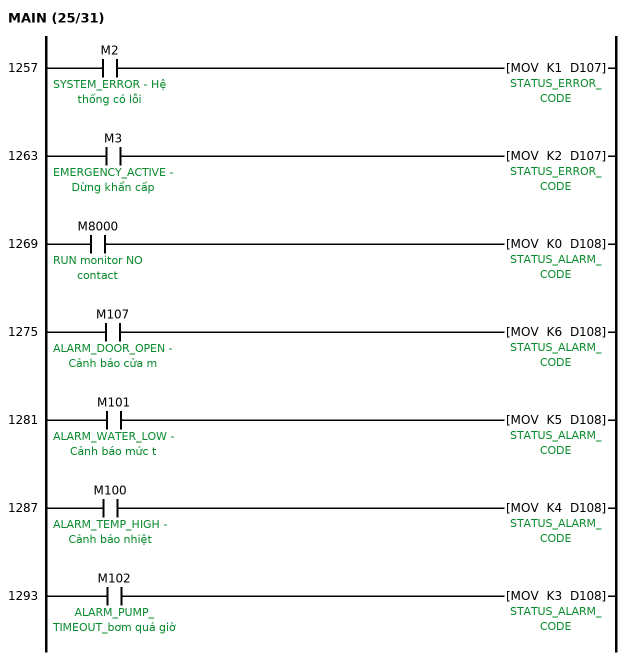
[picture p24: ladder of MAIN, rungs at steps 1257 to 1293]
1257  LD      M2  ; SYSTEM_ERROR - Hệ thống có lỗi
      MOV     K1 D107
1263  LD      M3  ; EMERGENCY_ACTIVE - Dừng khẩn cấp
      MOV     K2 D107
1269  LD      M8000  ; RUN monitor NO contact
      MOV     K0 D108  ; STATUS_ALARM_CODE
1275  LD      M107  ; ALARM_DOOR_OPEN - Cảnh báo cửa m
      MOV     K6 D108
1281  LD      M101  ; ALARM_WATER_LOW - Cảnh báo mức t
      MOV     K5 D108
1287  LD      M100  ; ALARM_TEMP_HIGH - Cảnh báo nhiệt
      MOV     K4 D108
1293  LD      M102  ; ALARM_PUMP_TIMEOUT_bơm quá giờ
      MOV     K3 D108
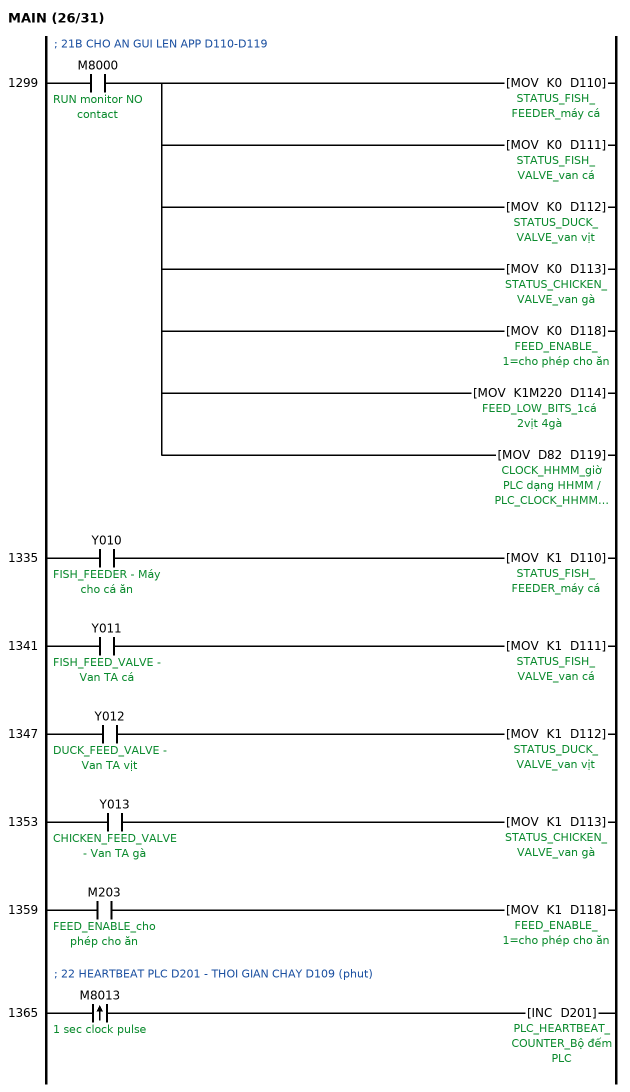
; 21B CHO AN GUI LEN APP D110-D119
1299  LD      M8000  ; RUN monitor NO contact
      MOV     K0 D110  ; STATUS_FISH_FEEDER_máy cá
      MOV     K0 D111  ; STATUS_FISH_VALVE_van cá
      MOV     K0 D112  ; STATUS_DUCK_VALVE_van vịt
      MOV     K0 D113  ; STATUS_CHICKEN_VALVE_van gà
      MOV     K0 D118  ; FEED_ENABLE_1=cho phép cho ăn
      MOV     K1M220 D114  ; FEED_LOW_BITS_1cá 2vịt 4gà
      MOV     D82 D119  ; PLC_CLOCK_HHMM_giờ PLC
1335  LD      Y010  ; FISH_FEEDER - Máy cho cá ăn
      MOV     K1 D110
1341  LD      Y011  ; FISH_FEED_VALVE - Van TA cá
      MOV     K1 D111
1347  LD      Y012  ; DUCK_FEED_VALVE - Van TA vịt
      MOV     K1 D112
1353  LD      Y013  ; CHICKEN_FEED_VALVE - Van TA gà
      MOV     K1 D113
1359  LD      M203  ; FEED_ENABLE_cho phép cho ăn
      MOV     K1 D118
; 22 HEARTBEAT PLC D201 - THOI GIAN CHAY D109 (phut)
1365  LDP     M8013  ; 1 sec clock pulse
      INC     D201  ; PLC_HEARTBEAT_COUNTER_Bộ đếm PLC
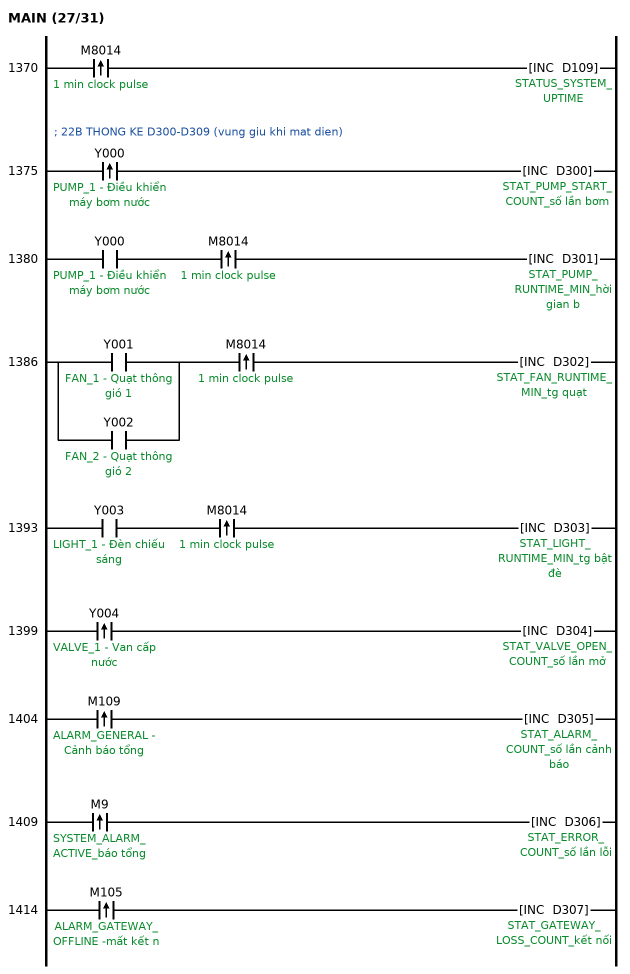
1370  LDP     M8014  ; 1 min clock pulse
      INC     D109  ; STATUS_SYSTEM_UPTIME
; 22B THONG KE D300-D309 (vung giu khi mat dien)
1375  LDP     Y000  ; PUMP_1 - Điều khiển máy bơm nước
      INC     D300  ; STAT_PUMP_START_COUNT_số lần bơm
1380  LD      Y000  ; PUMP_1 - Điều khiển máy bơm nước
      ANDP    M8014  ; 1 min clock pulse
      INC     D301  ; STAT_PUMP_RUNTIME_MIN_hời gian b
1386  LD      Y001  ; FAN_1 - Quạt thông gió 1
      OR      Y002  ; FAN_2 - Quạt thông gió 2
      ANDP    M8014  ; 1 min clock pulse
      INC     D302  ; STAT_FAN_RUNTIME_MIN_tg quạt
1393  LD      Y003  ; LIGHT_1 - Đèn chiếu sáng
      ANDP    M8014  ; 1 min clock pulse
      INC     D303  ; STAT_LIGHT_RUNTIME_MIN_tg bật đè
1399  LDP     Y004  ; VALVE_1 - Van cấp nước
      INC     D304  ; STAT_VALVE_OPEN_COUNT_số lần mở
1404  LDP     M109  ; ALARM_GENERAL - Cảnh báo tổng
      INC     D305  ; STAT_ALARM_COUNT_số lần cảnh báo
1409  LDP     M9  ; SYSTEM_ALARM_ACTIVE_báo tổng
      INC     D306  ; STAT_ERROR_COUNT_số lần lỗi
1414  LDP     M105  ; ALARM_GATEWAY_OFFLINE -mất kết n
      INC     D307  ; STAT_GATEWAY_LOSS_COUNT_kết nối
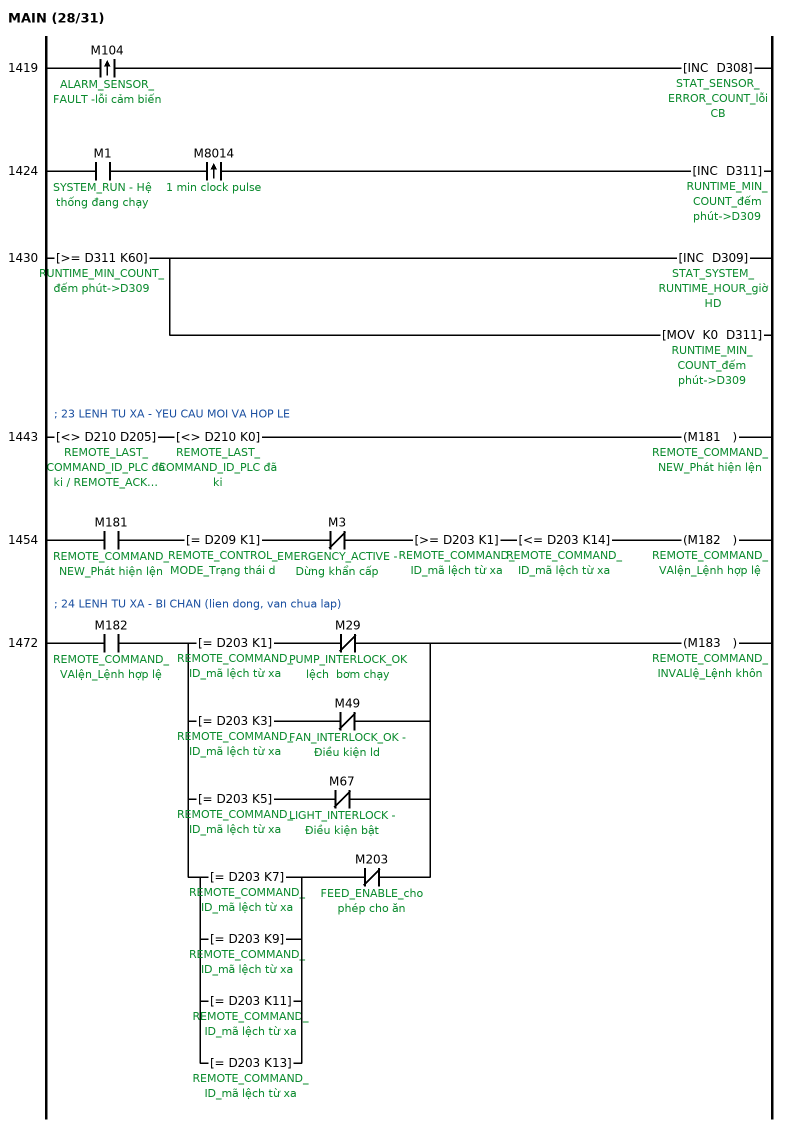
1419  LDP     M104  ; ALARM_SENSOR_FAULT -lỗi cảm biến
      INC     D308  ; STAT_SENSOR_ERROR_COUNT_lỗi CB
1424  LD      M1  ; SYSTEM_RUN - Hệ thống đang chạy
      ANDP    M8014  ; 1 min clock pulse
      INC     D311  ; RUNTIME_MIN_COUNT_đếm phút->D309
1430  LD>=    D311 K60  ; RUNTIME_MIN_COUNT_đếm phút->D309
      INC     D309  ; STAT_SYSTEM_RUNTIME_HOUR_giờ HD
      MOV     K0 D311
; 23 LENH TU XA - YEU CAU MOI VA HOP LE
1443  LD<>    D210 D205  ; REMOTE_LAST_COMMAND_ID_PLC đã ki / REMOTE_ACK_COMMAND_ID_PLC đã nhậ
      AND<>   D210 K0  ; REMOTE_LAST_COMMAND_ID_PLC đã ki
      OUT     M181  ; REMOTE_COMMAND_NEW_Phát hiện lện
1454  LD      M181  ; REMOTE_COMMAND_NEW_Phát hiện lện
      AND=    D209 K1  ; REMOTE_CONTROL_MODE_Trạng thái d
      ANI     M3  ; EMERGENCY_ACTIVE - Dừng khẩn cấp
      AND>=   D203 K1  ; REMOTE_COMMAND_ID_mã lệch từ xa
      AND<=   D203 K14  ; REMOTE_COMMAND_ID_mã lệch từ xa
      OUT     M182  ; REMOTE_COMMAND_VAlện_Lệnh hợp lệ
; 24 LENH TU XA - BI CHAN (lien dong, van chua lap)
1472  LD      M182  ; REMOTE_COMMAND_VAlện_Lệnh hợp lệ
      LD=     D203 K1  ; REMOTE_COMMAND_ID_mã lệch từ xa
      ANI     M29  ; PUMP_INTERLOCK_OK lệch  bơm chạy
      LD=     D203 K3  ; REMOTE_COMMAND_ID_mã lệch từ xa
      ANI     M49  ; FAN_INTERLOCK_OK - Điều kiện ld
      ORB
      LD=     D203 K5  ; REMOTE_COMMAND_ID_mã lệch từ xa
      ANI     M67  ; LIGHT_INTERLOCK - Điều kiện bật
      ORB
      LD=     D203 K7  ; REMOTE_COMMAND_ID_mã lệch từ xa
      OR=     D203 K9  ; REMOTE_COMMAND_ID_mã lệch từ xa
      OR=     D203 K11  ; REMOTE_COMMAND_ID_mã lệch từ xa
      OR=     D203 K13  ; REMOTE_COMMAND_ID_mã lệch từ xa
      ANI     M203  ; FEED_ENABLE_cho phép cho ăn
      ORB
      ANB
      OUT     M183  ; REMOTE_COMMAND_INVALlệ_Lệnh khôn
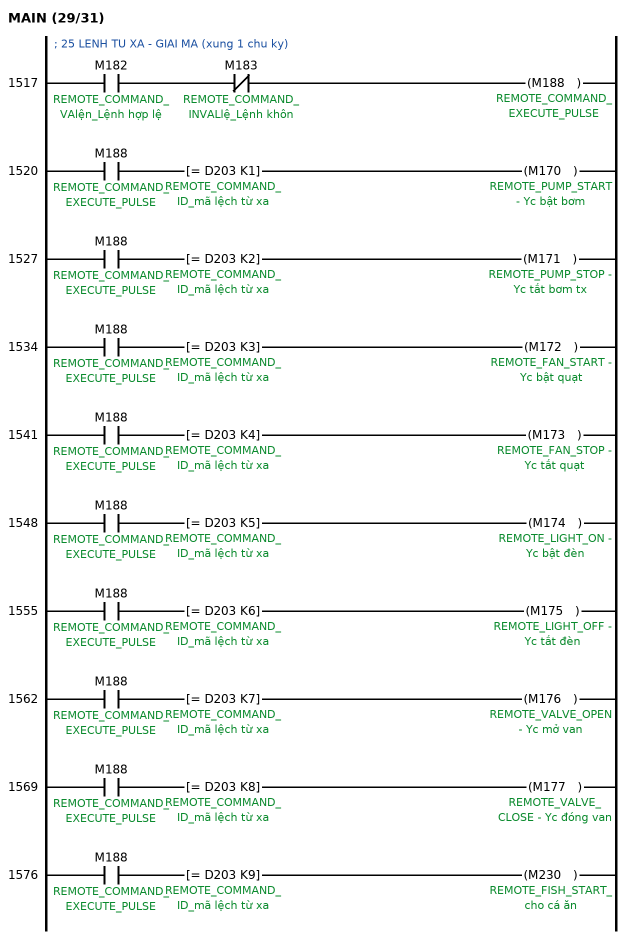
; 25 LENH TU XA - GIAI MA (xung 1 chu ky)
1517  LD      M182  ; REMOTE_COMMAND_VAlện_Lệnh hợp lệ
      ANI     M183  ; REMOTE_COMMAND_INVALlệ_Lệnh khôn
      OUT     M188  ; REMOTE_COMMAND_EXECUTE_PULSE
1520  LD      M188  ; REMOTE_COMMAND_EXECUTE_PULSE
      AND=    D203 K1  ; REMOTE_COMMAND_ID_mã lệch từ xa
      OUT     M170  ; REMOTE_PUMP_START - Yc bật bơm
1527  LD      M188  ; REMOTE_COMMAND_EXECUTE_PULSE
      AND=    D203 K2  ; REMOTE_COMMAND_ID_mã lệch từ xa
      OUT     M171  ; REMOTE_PUMP_STOP - Yc tắt bơm tx
1534  LD      M188  ; REMOTE_COMMAND_EXECUTE_PULSE
      AND=    D203 K3  ; REMOTE_COMMAND_ID_mã lệch từ xa
      OUT     M172  ; REMOTE_FAN_START - Yc bật quạt
1541  LD      M188  ; REMOTE_COMMAND_EXECUTE_PULSE
      AND=    D203 K4  ; REMOTE_COMMAND_ID_mã lệch từ xa
      OUT     M173  ; REMOTE_FAN_STOP - Yc tắt quạt
1548  LD      M188  ; REMOTE_COMMAND_EXECUTE_PULSE
      AND=    D203 K5  ; REMOTE_COMMAND_ID_mã lệch từ xa
      OUT     M174  ; REMOTE_LIGHT_ON - Yc bật đèn
1555  LD      M188  ; REMOTE_COMMAND_EXECUTE_PULSE
      AND=    D203 K6  ; REMOTE_COMMAND_ID_mã lệch từ xa
      OUT     M175  ; REMOTE_LIGHT_OFF - Yc tắt đèn
1562  LD      M188  ; REMOTE_COMMAND_EXECUTE_PULSE
      AND=    D203 K7  ; REMOTE_COMMAND_ID_mã lệch từ xa
      OUT     M176  ; REMOTE_VALVE_OPEN - Yc mở van
1569  LD      M188  ; REMOTE_COMMAND_EXECUTE_PULSE
      AND=    D203 K8  ; REMOTE_COMMAND_ID_mã lệch từ xa
      OUT     M177  ; REMOTE_VALVE_CLOSE - Yc đóng van
1576  LD      M188  ; REMOTE_COMMAND_EXECUTE_PULSE
      AND=    D203 K9  ; REMOTE_COMMAND_ID_mã lệch từ xa
      OUT     M230  ; REMOTE_FISH_START_cho cá ăn
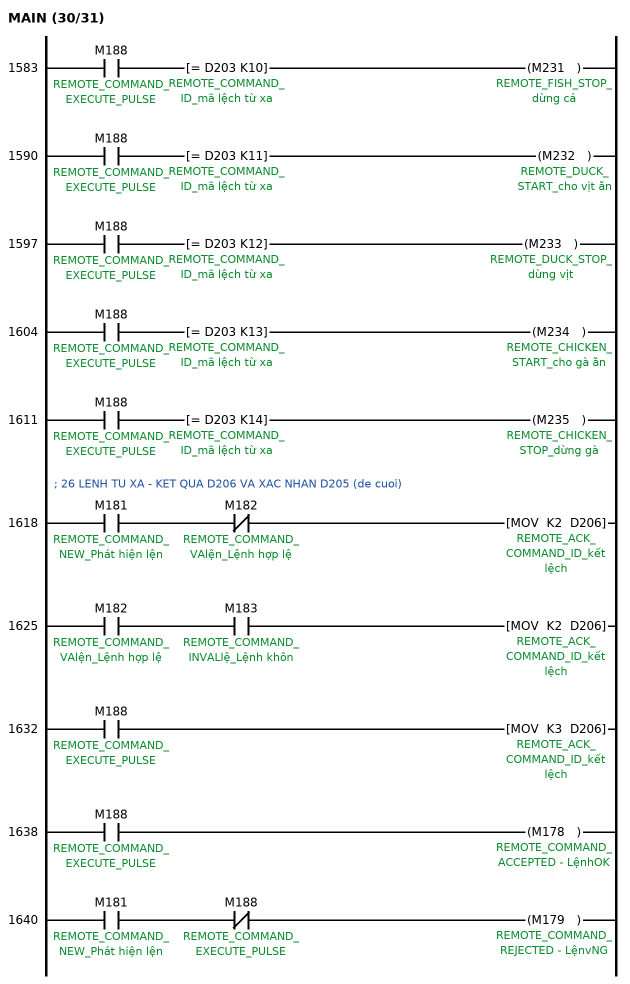
1583  LD      M188  ; REMOTE_COMMAND_EXECUTE_PULSE
      AND=    D203 K10  ; REMOTE_COMMAND_ID_mã lệch từ xa
      OUT     M231  ; REMOTE_FISH_STOP_dừng cá
1590  LD      M188  ; REMOTE_COMMAND_EXECUTE_PULSE
      AND=    D203 K11  ; REMOTE_COMMAND_ID_mã lệch từ xa
      OUT     M232  ; REMOTE_DUCK_START_cho vịt ăn
1597  LD      M188  ; REMOTE_COMMAND_EXECUTE_PULSE
      AND=    D203 K12  ; REMOTE_COMMAND_ID_mã lệch từ xa
      OUT     M233  ; REMOTE_DUCK_STOP_dừng vịt
1604  LD      M188  ; REMOTE_COMMAND_EXECUTE_PULSE
      AND=    D203 K13  ; REMOTE_COMMAND_ID_mã lệch từ xa
      OUT     M234  ; REMOTE_CHICKEN_START_cho gà ăn
1611  LD      M188  ; REMOTE_COMMAND_EXECUTE_PULSE
      AND=    D203 K14  ; REMOTE_COMMAND_ID_mã lệch từ xa
      OUT     M235  ; REMOTE_CHICKEN_STOP_dừng gà
; 26 LENH TU XA - KET QUA D206 VA XAC NHAN D205 (de cuoi)
1618  LD      M181  ; REMOTE_COMMAND_NEW_Phát hiện lện
      ANI     M182  ; REMOTE_COMMAND_VAlện_Lệnh hợp lệ
      MOV     K2 D206
1625  LD      M182  ; REMOTE_COMMAND_VAlện_Lệnh hợp lệ
      AND     M183  ; REMOTE_COMMAND_INVALlệ_Lệnh khôn
      MOV     K2 D206
1632  LD      M188  ; REMOTE_COMMAND_EXECUTE_PULSE
      MOV     K3 D206
1638  LD      M188  ; REMOTE_COMMAND_EXECUTE_PULSE
      OUT     M178  ; REMOTE_COMMAND_ACCEPTED - LệnhOK
1640  LD      M181  ; REMOTE_COMMAND_NEW_Phát hiện lện
      ANI     M188  ; REMOTE_COMMAND_EXECUTE_PULSE
      OUT     M179  ; REMOTE_COMMAND_REJECTED - LệnvNG
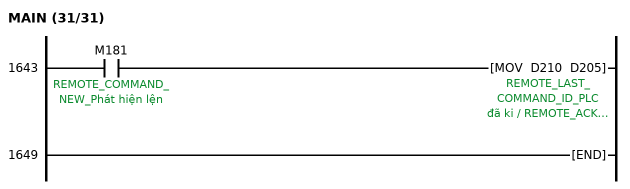
1643  LD      M181  ; REMOTE_COMMAND_NEW_Phát hiện lện
      MOV     D210 D205
1649  END
END_PROGRAM

// device comments not shown above
M7  ; AUTO_ENABLE - Cho phép chế độ tự
M8  ; MANUAL_ENABLE - Cho phép chế độ
M15  ; MODE_INITIALIZING_Trạng thái HT
M26  ; PUMP_FAULT - Lỗi máy bơm
M50  ; FAN_AUTO_RUN_LATCH_bit nhớ
M52  ; FAN2_AUTO_STATE_trạng thái bật/t
M54  ; FAN2_MANUAL_STATE_trạng thái bật
M66  ; LIGHT_FAULT - Lỗi hệ thống đèn
M80  ; VALVE_AUTO_REQUEST_mở tự động
M81  ; VALVE_MANUAL_REQUEST -mở thủ côn
M82  ; VALVE_REMOTE_REQUEST -mở từ xa
M84  ; VALVE_CLOSE_CMD - Lệnh đóng van
M85  ; VALVE_OPENING - Trạng thái mở
M86  ; VALVE_FAULT - Lỗi van cấp nước
M87  ; VALVE_INTERLOCK- Điều kiện mở
M88  ; WATER_SUPPLY_ACTIVE - Đang cấp n
M89  ; VALVE_TIMEOUT - Van hd quá giờ
M103  ; ALARM_FAN_FAULT - Cảnh báo quạt
M106  ; ALARM_WATER_HIGH - nước quá cao
M108  ; ALARM_POWER_FAIL - mất nguồn
M130  ; ERROR_TEMP_SENSOR - Lỗi cb nhiệt
M131  ; ERROR_HUMIDITY_SENSOR - Lỗi da
M133  ; ERROR_PUMP - Lỗi máy bơm
M134  ; ERROR_FAN - Lỗi quạt
M135  ; ERROR_VALVE - Lỗi van nước
M136  ; ERROR_GATEWAY - Lỗi Gateway
M137  ; ERROR_COMMUNICATION - Lỗi RS485
M138  ; ERROR_OVERLOAD - Lỗi quá tải thi
M139  ; ERROR_SYSTEM - Lỗi tổng hệ thống
M150  ; GATEWAY_ONLINE - Gateway kết nối
M151  ; GATEWAY_COMMAND_VALID - Lệnh OK
M152  ; GATEWAY_DATA_READY - Dữ liệu SS
M153  ; RS485_TX_REQUEST - gửi dữ liệu
M154  ; RS485_RX_COMPLETE - Nhận dữ liệu
M155  ; RS485_COMM_ERROR - Lỗi RS485
M156  ; PLC_HEARTBEAT - Xung kiểm traPLC
M157  ; GATEWAY_HEARTBEAT -kiểm tra gate
M158  ; COMM_TIMEOUT - Quá thời gian phả
M159  ; COMM_RECOVERY - Đã khôi phục kết
M184  ; REMOTE_COMMAND_PROCESkhôn_Đang x
M185  ; REMOTE_COMMAND_DONE_Đã xử lý xon
M186  ; REMOTE_COMMAND_Bxon_Đang bận xử
M187  ; REMOTE_COMMAND_RESET_Xóa trạng t
D10  ; SET_TEMP_ALARM_LOW_nhiệt độ thấ
D51  ; SENSOR_AIR_HUMIDITY_độ ẩm
D52  ; SENSOR_WATER_TEMP_nhiệt độ nước
D53  ; SENSOR_WATER_LEVEL_mực nước
D54  ; SENSOR_SOIL_HUMIDITY_độ ẩm đất
D55  ; SENSOR_LIGHT_VALUE_độ sáng
D56  ; SENSOR_CO2_VALUE_Nồng độ CO₂
D57  ; SENSOR_NH3_VALUE_Nồng độ NH₃
D59  ; SENSOR_DATA_STATUS_trạng thái dl
D63  ; TEMP_FAN2_ON_bật quạt 2
D64  ; TEMP_FAN2_OFF_tắt quạt 2
D66  ; FAN_AUTO_DELAY_Thời gian trễ
D67  ; FAN_CONTROL_MODE_Chế độ điều khi
D68  ; FAN1_RUNTIME_Thời gian hoạt động
D69  ; FAN2_RUNTIME_Thời gian hoạt động
D204  ; REMOTE_COMMAND_VALUE_giá trị DK
D207  ; COMM_ERROR_CODE_Mã lỗi truyền th
D208  ; COMM_DATA_COUNTER_Bộ đếm dữ liệu
